(* IEC 61131-3 sources: BODAS-HelloWorld/st/bodas_rc18_12_40/plc_logic/application/02_easyconfig/easyconfig_import/bds_sysio_ec, 6 files *)

(* ---- bds_sys_ait_signal_te-bds_sys_ait_signal_te.st ---- *)
(* --- Interface --- *)
{attribute 'qualified_only' := ''}
{attribute 'strict' := ''}
TYPE bds_sys_ait_signal_te : (
		SYS_AIT_START_SIGNALS := 16#900,
		SYS_AIT_START         := 16#8FF,
		TSGI1,
		TSGI2,
		SYS_AIT_NUM_SIGNALS
	) UINT;
END_TYPE

(* ---- bds_sys_aiv_signal_te-bds_sys_aiv_signal_te.st ---- *)
(* --- Interface --- *)
{attribute 'qualified_only' := ''}
{attribute 'strict' := ''}
TYPE bds_sys_aiv_signal_te : (
		SYS_AIV_START_SIGNALS := 16#A00,
		SYS_AIV_START         := 16#9FF,
		UBAT_MON,
		UBRM24_MON,
		VDD5A_MON,
		UBR24_VP,
		UBRM24_LOADS,
		VDD3V3,
		VPR6,
		VDD5V_IN,
		VDD5_S3530,
		VSS3V5,
		VSS4V10,
		LSS_MEAS_CL13,
		LSS_MEAS_CL2,
		SYS_AIV_NUM_SIGNALS
	) UINT;
END_TYPE

(* ---- bds_sys_di_signal_te-bds_sys_di_signal_te.st ---- *)
(* --- Interface --- *)
{attribute 'qualified_only' := ''}
{attribute 'strict' := ''}
TYPE bds_sys_di_signal_te : (
		SYS_DI_START_SIGNALS := 16#D00,
		SYS_DI_START         := 16#CFF,
		ST_INH,
		SYS_DI_NUM_SIGNALS
	) UINT;
END_TYPE

(* ---- bds_sys_do_signal_te-bds_sys_do_signal_te.st ---- *)
(* --- Interface --- *)
{attribute 'qualified_only' := ''}
{attribute 'strict' := ''}
TYPE bds_sys_do_signal_te : (
		SYS_DO_START_SIGNALS := 16#B00,
		SYS_DO_START         := 16#AFF,
		SHUNT_AIC_K39_EN,
		SHUNT_AIC_K38_EN,
		SHUNT_AIC_K40_EN,
		SHUNT_AIC_K41_EN,
		SHUNT_AIC_K42_EN,
		SHUNT_AIC_K45_EN,
		SHUNT_AIC_K44_EN,
		SHUNT_AIC_K65_EN,
		SHUNT_AIC_K63_EN,
		SHUNT_AIC_K64_EN,
		SHUNT_AIC_A36_EN,
		SHUNT_AIC_A37_EN,
		SHUNT_AIC_A38_EN,
		SHUNT_AIC_A39_EN,
		SHUNT1_EN,
		SHUNT3_EN,
		SHUNT5_EN,
		SHUNT6_EN,
		SYS_DO_NUM_SIGNALS
	) UINT;
END_TYPE

(* ---- bds_sys_vss_signal_te-bds_sys_vss_signal_te.st ---- *)
(* --- Interface --- *)
{attribute 'qualified_only' := ''}
{attribute 'strict' := ''}
TYPE bds_sys_vss_signal_te : (
		SYS_VSS_START_SIGNALS := 16#C00,
		SYS_VSS_START         := 16#BFF,
		VSS1,
		VSS2,
		VSS3,
		VSS4,
		SYS_VSS_NUM_SIGNALS,
		SYS_VSS_CY_NUM_SIGNALS := VSS3
	) UINT;
END_TYPE

(* ---- bds_sysio_ec_gvl-bds_sysIo_ec_gvl.st ---- *)
(* --- Interface --- *)
{attribute 'qualified_only' := ''}
VAR_GLOBAL CONSTANT
	BDS_SYSIO_FI_SHUNT_NUM_SIGNALS_D : UINT := bds_sys_do_signal_te.SHUNT1_EN;
END_VAR
